// Communication API/ISOBUS/J1939-76/API/bds_isobus_initCnsrSdgDatabox
///This function initializes a J1939-76 consumer databox. The  J1939-76 messages can be sent only with  J1939-76 consumer databoxes.
///
///=======
/// Remarks:
///=======
/// + This function must be called during the configuration of the ISOBUS/J1939 and J1939-76 communication stack once for each J1939-76 consumer message.
/// + Before the consumer databoxes can be initialized with this function, the required number of receive databoxes has to be configured first with easyConfig tool or alternatively with function bds_isobus_registerCnsrSdgDataboxes.
/// + Each J1939-76 consumer databox requires an own data array or a data structure. The pointer to this data field is required for the initialization of a J1939-76 consumer databox. The received data then will be stored in this data field.
/// + The data array for the received data shall have length less than or equal to 8 (see parameter description below). 
/// + The execution time of the callback function should be short to be able to meet the time conditions within the ISOBUS/J1939 stack.
/// + If the same CAN bus is also used for further communication, ensure that the CAN IDs are uniquely assigned.
/// + The meaning of this function is similar to the ISOBUS/J1939 function bds_isobus_initRxDatabox.
/// + In addition to the ISOBUS/J1939 specifications, this function can be used for the reception of J1939-76 PDU1 format messages which are sent to the own network adddress as well as to other destination addresses.
/// + The definition of a destination address within PDU1 format PGNs is mandatory.
/// + Important: For the reception of PDU1 format messages to the own network address the PDU specific part (=Destination) of the PGN should be defined with the NULL address value (=0xFE) instead of the own address. Otherwise the own address within the RX databoxes may not match any more with the real own address after an address claiming.  
/// + The header file bds_bsw.h is included for enabling usage of defines.
///
///----------
/// FFI:
///----------
///This API can be used in trusted partitions only. See Freedom from Interference (FFI) concept for more details.
///
///
///Return value    																		Description
///==================================================================		  			===================================================================================================
///0: bds_isobus_sfty_noErr_E															Function executed without error
///3: bds_isobus_sfty_invldInstNum_E													Invalid ISOBUS/J1939 CA instance number
///7: bds_isobus_sfty_invldDataboxNum_E													Invalid databox number
///8: bds_isobus_sfty_invldPgn_E														Invalid PGN
///9: bds_isobus_sfty_invldPrio_E														Invalid priority
///10: bds_isobus_sfty_invldCyc_E														Invalid cycle time
///11: bds_isobus_sfty_invldOffs_E														Invalid offset time.
///12: bds_isobus_sfty_invldDataLen_E													Invalid data length
///13: bds_isobus_sfty_invldDataPtr_E													invalid pointer address
///14: bds_isobus_sfty_pgnPrioExists_E													Another databox with the same PGN and priority is already defined.
///15: bds_isobus_sfty_invldSrcAdr_E													Invalid Source Address
///16: bds_isobus_sfty_invldSct_E														Invalid SCT value
///17: bds_isobus_sfty_invldSrvt_E														Invalid SRVT value	
///19: bds_isobus_sfty_featNotEnad_E													API used without enabling J1939-76 feature in easyConfig
///20: bds_isobus_sfty_invldCbkAdr_E 													Callback function value NULL is invalid. Callback function is mandatory for J1939-76
///					  									
///==================================================================		   			===================================================================================================
///
///
///==================================================================		  			===================================================================================================
///Standard PGN	 								  										Data in Databox
///==================================================================		  			===================================================================================================
///Registered as "0xEEFF"																Receives only data which is broadcasted (PDU Specific part =0xFF).
///																						ex: bds_isobus_initCnsrSdgDatabox(1u, 1u, 0xEEFF, 0x10, 120, 50, 8, cnsrSDMdata_au8, NULL);
///																						It only receives the data which is brodcasted from source address 0x10.
///
///Registered "0xEE<own address>"														Receives data which is directed to the ECU by its own address (PDU Specific part=Destination).
///																						ex: bds_isobus_initCnsrSdgDatabox(1u, 1u, 0xEE04, 0x10, 120, 50, 8, cnsrSDMdata_au8, NULL);
///																						It only receives the data which is directed TO the ECU BY requesting with its own address(0x04).
///																					    Note: IF you initialize databox with "0xEEFE" you only receive data with whose PDU Specific part is Null(0xFE).
///==================================================================		   			===================================================================================================
///
///=======
///Code Example:
///=======
///============================================================================
///
/// PROGRAM Isobus_test
/// VAR_GLOBAL
///  cnsrMsg1Data_au8: ARRAY[1..8] OF USINT;
///
/// END_VAR
///	
/// 
/// VAR
///	   ISOBUS_SFTY_CNSR_BOXES_DU8: USINT :=35;
///    registerApiRetVal_e : bds_isobus_sfty_apiRetVal_te;    
///    initApi1RetVal_e : bds_isobus_sfty_apiRetVal_te;
///    isobus_sfty_cnsrSdgMsg_as: ARRAY[1..35] OF bds_isobus_cnsrSdgMsg_ts ;
///    instance_num:USINT:=1;
///
/// END_VAR
///
/// IF(Flag_u8=0) THEN
///
/// bds_can_init(BDS_CAN_3_D, BDS_BAUD_1000K_DU32); 	
///	bds_can_sendData(BDS_CAN_3_D, 16#999999, 1, 0,0);
///
/// registerApiRetVal_e := bds_isobus_registerCnsrSdgDataboxes(1, ADR(isobus_sfty_cnsrSdgMsg_as), ISOBUS_SFTY_CNSR_BOXES_DU8);
/// 
/// initApi1RetVal_e := bds_isobus_initCnsrSdgDatabox(1, 1, 16#4901, 16#10, 24, 100, 8, ADR(gvl.cnsrMsg1Data_au8), ADR(cnsrMsgCallback1));
///
/// bds_isobus_setCaName(instance_num,16#00,16#02,16#00,16#01,16#81,16#01,16#01,16#33,BDS_ISOBUS_OWN_SN_DU32);
///
/// bds_isobus_setCaName(instance_num,16#00,16#02,16#00,16#01,16#81,16#01,16#01,16#33,BDS_ISOBUS_OWN_SN_DU32);
/// 
/// retval5_u16:=bds_isobus_setCaAddr(instance_num,BDS_CAN_3_D,16#10);
///
/// bds_isobus_initComm(bds_can_Chnl_te.BDS_CAN_3_D, 50);
///
/// Flag_u8:=1;
/// 
/// END_IF
///
/// FUNCTION cnsrMsgCallback1 : UINT
/// VAR_INPUT	
///	data_length: POINTER TO BYTE;
///	data_pau8: POINTER TO BYTE ;
///	status_e : bds_isobus_sdgCnsrStatus_te;
/// END_VAR

/// VAR
///  i : INT;
///    cnsrCbk_rcvd_u32 : UDINT;
///    CbkSt_e : bds_isobus_sdgCnsrStatus_te;
///    CbkDataLen_u8 : POINTER TO BYTE:=0;
///	 data_au8: ARRAY [1..8] OF USINT:=[1,2];
/// END_VAR
///
/// cnsrCbk_rcvd_u32 := cnsrCbk_rcvd_u32 + 1;
/// CbkDataLen_u8 := data_length;
/// CbkSt_e := status_e;
///
/// FOR i := 0 TO 7 DO
/// gvl.cnsrMsg1Data_au8[i] := data_pau8[i];  // Dereference pointer to copy each element
/// END_FOR;
/// END
///============================================================================

{attribute 'external_name' := 'cmp_rts_bds_isobus_initCnsrSdgDatabox'}

FUNCTION bds_isobus_initCnsrSdgDatabox : bds_isobus_sfty_apiRetVal_te
VAR_INPUT
	///ISOBUS/J1939 instance number. This number identifies one instance of the ISOBUS/J1939 stack.
 	///
	///Value range: 1..n
	///n is the number of ISOBUS instances configured by easyConfig. 
	instanceNum_u8 : USINT;
	///Number of a J1939-76 producer databox.
	///
	///Value range: 1..n
	///n is the number of producer databoxes configured by easyConfig or alternatively with function bds_isobus_registerProdSdgDataboxes.
	sdgDataboxNum_u16 : UINT;
	///Parameter group number (PGN) of the SDM(Safety Data Message) to be sent with this databox.
	///
	///Value range: 0..0x3FFFF (18 bit) 
	///The lowest byte of the PGN contains for:
	/// + PDU1 format:  the destination address
	/// + PDU2 format:  the PDU extension
	pgn_u32 : UDINT;
	///Source address of the J1939-76 consumer from where the message has to be received.
	///
	///
	///Value range: 0x00..0xFD 
	src_u8 : USINT;
	///The maximum time interval in ms between two consecutive SDMs received.
	///
	///
	///Value Range: 10ms - 65000ms
	sct_u32 : UDINT;
	///The maximum time interval in ms between an SHM and SDM of an SDG received.
	///
	///
	///Value Range: 10ms - 65000ms
	srvt_u32 : UDINT;
	///Size of the data to be received. A J1939-76 consumer message data size must be less than or equal to 8 bytes.
	//
	///Value range: 1...8 bytes
	lenMax_u8 : USINT;
	///Pointer to a data array, in which the received data can be stored.
	/// The size of this array/structure has to be given within the previous parameter (lenMax_u8).
	///
	///It is neccessary to declare the data buffer array as a global variable.
	data_pau8: POINTER TO USINT;
	///Pointer to callback function of type bds_isobus_sdgCnsrCallback_tpf which will be called after reception and processing of a consumer SDG.
	func_pf: POINTER TO UINT;
END_VAR

END_FUNCTION

// Communication API/ISOBUS/J1939-76/API/bds_isobus_registerCnsrSdgDataboxes
///This function registers memory for J1939-76 safety extension consumer databoxes and therefore defines the maximal number of usable J1939-76 consumer databoxes per instance.
///
///=======
/// Remarks:
///=======
///		+ This function must be called once during the configuration of the ISOBUS/J1939 communication stack before bds_isobus_initComm.
/// 	+ After the execution of this function, each  J1939-76 consumer databox has to be initialized with bds_isobus_initCnsrSdgDatabox before using the databoxes.
/// 	+ The header file bds_bsw.h is included for enabling usage of defines.
/// 
///----------
/// FFI:
///----------
///
///This API can be used in trusted partitions only. See Freedom from Interference (FFI) concept for more details.
///	
///==================================================================		  			===================================================================================================
///Return value    								  									Description
///==================================================================		  			===================================================================================================
/// 0: bds_isobus_sfty_noErr_E 																Function executed without error
/// 1: bds_isobus_sfty_invldAdr_E															invalid address of databox (mem_pas)
/// 2: bds_isobus_sfty_ovlAdr_E                                                             Address overlaps with an already existing buffer.
/// 3: bds_isobus_sfty_invldInstNum_E                                                       Invalid CA instance number
///	6: bds_isobus_sfty_cfgNotAllwd_E                                                        Function must be called before bds_isobus_initComm, but it was called afterwards.																			-
/// 19: bds_isobus_sfty_featNotEnad_E                                                       API used without enabling J1939-76 feature in easyConfig
///
///
///==================================================================		   			===================================================================================================
///
/// Code Example:
///=======
///============================================================================
/// PROGRAM Isobus_test
/// VAR_GLOBAL
///  cnsrMsg1Data_au8: ARRAY[1..8] OF USINT;
///
/// END_VAR
///	
/// 
/// VAR
///	   ISOBUS_SFTY_CNSR_BOXES_DU8: USINT :=35;
///    registerApiRetVal_e : bds_isobus_sfty_apiRetVal_te;    
///    initApi1RetVal_e : bds_isobus_sfty_apiRetVal_te;
///    isobus_sfty_cnsrSdgMsg_as: ARRAY[1..35] OF bds_isobus_cnsrSdgMsg_ts ;
///    instance_num:USINT:=1;
///
/// END_VAR
///
/// IF(Flag_u8=0) THEN
///
/// bds_can_init(BDS_CAN_3_D, BDS_BAUD_1000K_DU32); 	
///	bds_can_sendData(BDS_CAN_3_D, 16#999999, 1, 0,0);
///
/// registerApiRetVal_e := bds_isobus_registerCnsrSdgDataboxes(1, ADR(isobus_sfty_cnsrSdgMsg_as), ISOBUS_SFTY_CNSR_BOXES_DU8);
/// 
/// initApi1RetVal_e := bds_isobus_initCnsrSdgDatabox(1, 1, 16#4901, 16#10, 24, 100, 8, ADR(gvl.cnsrMsg1Data_au8), ADR(cnsrMsgCallback1));
///
/// bds_isobus_setCaName(instance_num,16#00,16#02,16#00,16#01,16#81,16#01,16#01,16#33,BDS_ISOBUS_OWN_SN_DU32);
///
/// bds_isobus_setCaName(instance_num,16#00,16#02,16#00,16#01,16#81,16#01,16#01,16#33,BDS_ISOBUS_OWN_SN_DU32);
/// 
/// retval5_u16:=bds_isobus_setCaAddr(instance_num,BDS_CAN_3_D,16#10);
///
/// bds_isobus_initComm(bds_can_Chnl_te.BDS_CAN_3_D, 50);
///
/// Flag_u8:=1;
/// 
/// END_IF
///
/// FUNCTION cnsrMsgCallback1 : UINT
/// VAR_INPUT	
///	data_length: POINTER TO BYTE;
///	data_pau8: POINTER TO BYTE ;
///	status_e : bds_isobus_sdgCnsrStatus_te;
/// END_VAR

/// VAR
///  i : INT;
///    cnsrCbk_rcvd_u32 : UDINT;
///    CbkSt_e : bds_isobus_sdgCnsrStatus_te;
///    CbkDataLen_u8 : POINTER TO BYTE:=0;
///	 data_au8: ARRAY [1..8] OF USINT:=[1,2];
/// END_VAR
///
/// cnsrCbk_rcvd_u32 := cnsrCbk_rcvd_u32 + 1;
/// CbkDataLen_u8 := data_length;
/// CbkSt_e := status_e;
///
/// FOR i := 0 TO 7 DO
/// gvl.cnsrMsg1Data_au8[i] := data_pau8[i];  // Dereference pointer to copy each element
/// END_FOR;
/// END
///============================================================================


{attribute 'external_name' := 'cmp_rts_bds_isobus_registerCnsrSdgDataboxes'}
FUNCTION bds_isobus_registerCnsrSdgDataboxes : bds_isobus_sfty_apiRetVal_te
VAR_INPUT
	///ISOBUS/J1939 instance number. This number identifies one instance of the ISOBUS/J1939 stack.
	///
	///Value range: 1..n
	///n is the number of ISOBUS/J1939 instances configured in easyConfig. 
	instanceNum_u8 : USINT;
	///Pointer to an array of data type bds_isobus_cnsrSdgMsg_ts.
	///
	///Note:
	///The buffer will be managed by the C-API. The application has only to declare the buffer (memory space).It is necessary to declare the buffer array as a global variable.
	mem_pas : POINTER TO  bds_isobus_prodSdgMsg_ts;
	///Size of the array above, which corresponds to the number of usable J1939-76 consumer databoxes.
	numOfMsg_u16: UINT;
END_VAR

END_FUNCTION

// Communication API/ISOBUS/J1939-76/API/bds_isobus_registerProdSdgDataboxes
///This function registers memory for J1939-76 safety extension producer databoxes and therefore defines the maximal number of usable J1939-76 producer databoxes per instance.
///
///=======
/// Remarks:
///=======
///		+ This function must be called once during the configuration of the ISOBUS/J1939 communication stack before bds_isobus_initComm.
/// 	+ After the execution of this function, each J1939-76 producer databox has to be initialized with bds_isobus_initProdDatabox before using the databoxes.
///     + The header file bds_bsw.h is included for enabling usage of defines.
///
///----------
/// FFI:
///----------
///This API can be used in trusted partitions only. See Freedom from Interference (FFI) concept for more details.
///
///==================================================================		  			===================================================================================================
///Return value    								  									     Description
///==================================================================		  			===================================================================================================
///0: bds_isobus_sfty_noErr_E															Function executed without error
///1: bds_isobus_sfty_invldAdr_E														Invalid address of databox (*mem_pas)
///2: bds_isobus_sfty_ovlAdr_E															Address overlaps with an already existing buffer.
///3: bds_isobus_sfty_invldInstNum_E													invalid CA instance number.
///6: bds_isobus_sfty_cfgNotAllwd_E														Function must be called before bds_isobus_initComm, but it was called afterwards.
///19: bds_isobus_sfty_featNotEnad_E													API used without enabling J1939-76 feature in easyConfig
///
/// 
///==================================================================		   			===================================================================================================
///
/// Code Example:
///=======
///============================================================================
/// PROGRAM Isobus_test
/// VAR_GLOBAL
///  prodMsg2Data_au8: ARRAY[1..8] OF USINT:=[16#A,16#1,16#2,16#3,16#4,16#5,16#6,16#7];
///
/// END_VAR
///
/// VAR
///
///    registerApiRetVal_e : bds_isobus_sfty_apiRetVal_te;    
///    initApi1RetVal_e : bds_isobus_sfty_apiRetVal_te;
///    isobus_sfty_prodSdgMsg_as: ARRAY[1..34] OF bds_isobus_prodSdgMsg_ts  ;
///    instance_num:USINT:=1;
///
/// END_VAR
///
/// IF(Flag_u8=0) THEN
///
/// bds_can_init(BDS_CAN_3_D, BDS_BAUD_1000K_DU32); 	
///	bds_can_sendData(BDS_CAN_3_D, 16#999999, 1, 0,0);
///
/// registerApiRetVal_e := bds_isobus_registerProdSdgDataboxes(instance_num,ADR(isobus_sfty_prodSdgMsg_as), 35);
/// 
/// initApi1RetVal_e := bds_isobus_initProdSdgDatabox(instance_num,1,16#4410,6, 100 , 10 , 8 , ADR(gvl.prodMsg2Data_au8) ,ADR(ProdMsgCallback1));
///
/// bds_isobus_setCaName(instance_num,16#00,16#02,16#00,16#01,16#81,16#01,16#01,16#33,BDS_ISOBUS_OWN_SN_DU32);
///
/// bds_isobus_setCaName(instance_num,16#00,16#02,16#00,16#01,16#81,16#01,16#01,16#33,BDS_ISOBUS_OWN_SN_DU32);
/// 
/// retval5_u16:=bds_isobus_setCaAddr(instance_num,BDS_CAN_3_D,16#10);
///
/// bds_isobus_initComm(bds_can_Chnl_te.BDS_CAN_3_D, 50);
///
/// Flag_u8:=1;
/// 
/// END_IF
///
/// FUNCTION ProdMsgCallback1 : USINT
/// 
/// VAR_INPUT
/// data_length:POINTER TO BYTE;
/// data_pau8: POINTER TO BYTE;
/// END_VAR
///
/// data_pau8[0] := 16#07;
/// data_pau8[1] := 16#06;
/// data_pau8[2] := 16#05;
/// data_pau8[3] := 16#04;
/// data_pau8[4] := 16#03;
/// data_pau8[5] := 16#FF;
/// data_pau8[6] := 16#FF;
/// data_pau8[7] := 16#FF;
/// 
/// data_length[0]:=8;
///
/// END
///============================================================================
{attribute 'external_name' := 'cmp_rts_bds_isobus_registerProdSdgDataboxes'}
FUNCTION bds_isobus_registerProdSdgDataboxes : bds_isobus_sfty_apiRetVal_te
VAR_INPUT
	///ISOBUS/J1939 instance number. This number identifies one instance of the ISOBUS/J1939 stack.
	///
	///Value range: 1..n
	///n is the number of ISOBUS/J1939 instances configured in easyConfig. 
	instanceNum_u8 : USINT;
	///Pointer to an array of data type bds_isobus_prodSdgMsg_ts. 
	///
	///Note:
	///The buffer will be managed by the C-API. The application has only to declare the buffer (memory space).
	///It is necessary to declare the buffer array as a global variable.
	mem_pas : POINTER TO  bds_isobus_prodSdgMsg_ts;
	///Size of the array, which corresponds to the number of usable J1939-76 producer databoxes.  
	numOfMsg_u16: UINT;
END_VAR

END_FUNCTION

// Communication API/ISOBUS/J1939-76/API/bds_isobus_initProdSdgDatabox
///This function initializes a J1939-76 producer databox. The J1939-76 messages can be sent only with J1939-76 producer databoxes.
///=======
/// Remarks:
///=======
/// + This function must be called during the configuration of the ISOBUS/J1939 and J1939-76 communication stack once for each J1939-76 producer message.
/// + Before the producer databoxes can be initialized with this function, the required number of producer databoxes has to be configured first with easyConfig tool or alternatively with function bds_isobus_registerProdSdgDataboxes.
/// + Each J1939-76 producer databox requires an own data array or a data structure. The pointer to this data field is required for the initialization of a J1939-76 producer databox. The transmitted data will be taken from this data field.
/// + The data array for the transmitted data must have a length of less than or equal to 8 bytes (see parameter description below).
/// + The execution time of the callback function should be short to be able to meet the time conditions within the ISOBUS/J1939 stack. 
/// + If the same CAN bus is also used for further communication, ensure that the CAN IDs are uniquely assigned.
/// + The meaning of this function is similar to the ISOBUS/J1939 function bds_isobus_initTxDatabox.
/// + The header file bds_bsw.h is included for enabling usage of defines.

///----------
/// FFI:
///----------
///This API can be used in trusted partitions only. See Freedom from Interference (FFI) concept for more details.
///
///==================================================================		  			===================================================================================================
///Return value    								  									Description
///==================================================================		  			===================================================================================================
///0: bds_isobus_sfty_noErr_E                                                             Function executed without error
///3: bds_isobus_sfty_invldInstNum_E                                                      Invalid ISOBUS/J1939 CA instance number
///7: bds_isobus_sfty_invldDataboxNum_E                                                   invalid databox number
///8: bds_isobus_sfty_invldPgn_E                                                          Invalid PGN
///9: bds_isobus_sfty_invldPrio_E                                                         Invalid priority
///10: bds_isobus_sfty_invldCyc_E                                                         Invalid cycle time
///11: bds_isobus_sfty_invldOffs_E                                                        Invalid offset time.
///12: bds_isobus_sfty_invldDataLen_E                                                     Invalid data length. 
///13: bds_isobus_sfty_invldDataPtr_E                                                     Invalid pointer address
///14: bds_isobus_sfty_pgnPrioExists_E                                                    Another databox with the same PGN and priority is already defined.

///==================================================================		   			===================================================================================================
///
///=======
///Code Example:
///=======
///
/// PROGRAM Isobus_test
/// VAR_GLOBAL
///  prodMsg2Data_au8: ARRAY[1..8] OF USINT:=[16#A,16#1,16#2,16#3,16#4,16#5,16#6,16#7];
///
/// END_VAR
///
/// VAR
///
///    registerApiRetVal_e : bds_isobus_sfty_apiRetVal_te;    
///    initApi1RetVal_e : bds_isobus_sfty_apiRetVal_te;
///    isobus_sfty_prodSdgMsg_as: ARRAY[1..34] OF bds_isobus_prodSdgMsg_ts  ;
///    instance_num:USINT:=1;
///
/// END_VAR
///
/// IF(Flag_u8=0) THEN
///
/// bds_can_init(BDS_CAN_3_D, BDS_BAUD_1000K_DU32); 	
///	bds_can_sendData(BDS_CAN_3_D, 16#999999, 1, 0,0);
///
/// registerApiRetVal_e := bds_isobus_registerProdSdgDataboxes(instance_num,ADR(isobus_sfty_prodSdgMsg_as), 35);
/// 
/// initApi1RetVal_e := bds_isobus_initProdSdgDatabox(instance_num,1,16#4410,6, 100 , 10 , 8 , ADR(gvl.prodMsg2Data_au8) ,ADR(ProdMsgCallback1));
///
/// bds_isobus_setCaName(instance_num,16#00,16#02,16#00,16#01,16#81,16#01,16#01,16#33,BDS_ISOBUS_OWN_SN_DU32);
///
/// bds_isobus_setCaName(instance_num,16#00,16#02,16#00,16#01,16#81,16#01,16#01,16#33,BDS_ISOBUS_OWN_SN_DU32);
/// 
/// retval5_u16:=bds_isobus_setCaAddr(instance_num,BDS_CAN_3_D,16#10);
///
/// bds_isobus_initComm(bds_can_Chnl_te.BDS_CAN_3_D, 50);
///
/// Flag_u8:=1;
/// 
/// END_IF
///
///
/// FUNCTION ProdMsgCallback1 : USINT
/// 
/// VAR_INPUT
/// data_length:POINTER TO BYTE;
/// data_pau8: POINTER TO BYTE;
/// END_VAR
///
/// data_pau8[0] := 16#07;
/// data_pau8[1] := 16#06;
/// data_pau8[2] := 16#05;
/// data_pau8[3] := 16#04;
/// data_pau8[4] := 16#03;
/// data_pau8[5] := 16#FF;
/// data_pau8[6] := 16#FF;
/// data_pau8[7] := 16#FF;
/// 
/// data_length[0]:=8;
///
/// END
///============================================================================

{attribute 'external_name' := 'cmp_rts_bds_isobus_initProdSdgDatabox'}
FUNCTION bds_isobus_initProdSdgDatabox : bds_isobus_sfty_apiRetVal_te
VAR_INPUT
	///ISOBUS/J1939 instance number. This number identifies one instance of the ISOBUS/J1939 stack.
 	///
	///Value range: 1..n
	///n is the number of ISOBUS instances configured by easyConfig. 
	instanceNum_u8 : USINT;
	///Number of a J1939-76 producer databox.
	///
	///Value range: 1..n
	///n is the number of producer databoxes configured by easyConfig or alternatively with function bds_isobus_registerProdSdgDataboxes.
	sdgDataboxNum_u16 : UINT;
	///Parameter group number (PGN) of the SDM(Safety Data Message) to be sent with this databox.
	///
	///Value range: 0..0x3FFFF (18 bit) 
	///The lowest byte of the PGN contains for:
	/// + PDU1 format:  the destination address
	/// + PDU2 format:  the PDU extension
	pgn_u32 : UDINT;
	///Priority of the message to be sent.
	///
	///Value range: 0..7  (6 = default value according ISOBUS/J1939 specification)
	prio_u8 : USINT;
	/// This time (in ms) controls the cyclic transmission (or) fixed transmission of the J1939-76 Producer message from this J1939-76 producer databox.
	///The cycle time of a J1939-76 producer message must be greater than or equal to 10ms.
	///Cycle time value 0 is invalid.
	///Value range: 10..65000 [ms].
	cycle_u16 : UINT;
	///The first transmission cycle of a J1939-76 producer message can be shortened by this offset time (in ms). 
	///This can be used to prevent CAN bus overload, if several messages have to be sent with the same cycle time.
	///With an offset = 0 the first message will be sent after the cycle time.
	///
	///Value range: 0.. (cycle_u16 - 1) [ms]
	offset_u16 : UINT;
	///Size of the data to be transmitted in bytes. A J1939-76 producer message data size must be less than or equal to 8.
	/// 
	///Value range: 1...8 bytes
	lenMax_u8 : USINT;
	///Pointer to a data array, from which the data is taken for transmission.  
	///The size of this array has to be given within the previous parameter (lenMax_u8).
	///
	///It is necessary to declare the data array as a global variable.
	data_pau8: POINTER TO USINT;
	///Pointer to callback function of type bds_isobus_sdgProdCallback_tpf which will be called by
	///BSW FOR data update BY ASW before transmission OF a producer SDG.
	func_pf: POINTER TO USINT;
END_VAR

END_FUNCTION

// Diagnostics API/UDS/API/Vehicle Identification Number(VIN) APIs/bds_uds_setVin
///This function sets the Vehicle Identification Number(VIN) of the ECU.
///
///=======
///Additional Info: + The Vehicle Identification Number(VIN) configured in the ECU is mapped to the DID 0xF190.
///					+ By default, the VIN has a value of B0DASMACH1NE00001.
///=======
///
///=======
/// Remarks: 
///=======
///			+ This function must be called from OsIniProc().
/// 		+ The header file bds_bsw.h is included for enabling usage of defines.
///
///-----------
///
/// FFI:
///----------
///This API can be used in trusted partitions only. See Freedom from Interference (FFI) concept for more details.
///
///
///==================================================================		  			===================================================================================================
///Return value    								  									Description
///==================================================================		  			===================================================================================================
///bds_udsCmn_ok_E																		API call successful.
///bds_udsCmn_invldPrm_E																API call invalid because of an invalid parameter.
///bds_udsCmn_outOfRng_E																Out of range, the array size should be less than or equal to 17 bytes.
///bds_udsCmn_notAvl_E																	not available (e.g. busy, called to early in init, system is in a mode that it cannot measure, etc)
///==================================================================		   			===================================================================================================
///
///=======
///Code Example:
///=======
///PROGRAM Vin_test
/// VAR
/// setVin_pau8:ARRAY[0..16] OF USINT:=[16#54,16#45 ,16#53 ,16#54 ,16#56 ,16#49 ,16#4E ,16#42 ,16#4F ,16#44 ,16#41 ,16#53 ,16#31 ,16#32 ,16#33 ,16#34 ,16#35];
/// flag_1:USINT;
/// retval_e:  bds_udsCmn_statusApi_te;
/// END_VAR
///
/// IF(flag_1=0) THEN
/// retval_e:=bds_uds_setVin(ADR(setVin_pau8),17);
/// flag_1:=1;
/// END_IF
//=============================================
{attribute 'external_name' := 'cmp_rts_bds_uds_setVin'}
FUNCTION bds_uds_setVin : bds_udsCmn_statusApi_te
VAR_INPUT
	//Pointer to set/configure the VIN data which is mapped to the DID 0xF190.
	data_pau8: POINTER TO USINT;
	//Size of the Vehicle Identification Number in bytes.
	size_u8: USINT;
END_VAR

END_FUNCTION

// Diagnostics API/UDS/API/Vehicle Identification Number(VIN) APIs/bds_uds_getVin
///This function reads the Vehicle Identification Number(VIN) of the ECU.
///
///=======
///Additional Info: + The Vehicle Identification Number(VIN) configured in the ECU is mapped to the DID 0xF190.
///					+ By default, the VIN has a value of B0DASMACH1NE00001.
///=======
///
///=======
/// Remarks: 
///=======
/// 		+ The header file bds_bsw.h is included for enabling usage of defines.
///
///-----------
///
/// FFI:
///----------
///This API can be used in trusted partitions only. See Freedom from Interference (FFI) concept for more details.
///
///
///==================================================================		  			===================================================================================================
///Return value    								  									Description
///==================================================================		  			===================================================================================================
///bds_udsCmn_ok_E																		API call successful.
///bds_udsCmn_invldPrm_E																API call invalid because of an invalid parameter.
///bds_udsCmn_outOfRng_E																Out of range, the array size should be less than or equal to 17 bytes.
///
///==================================================================		   			===================================================================================================
///
///=======
///Code Example:
///=======
///PROGRAM Vin_test
/// VAR
/// getVin_pau8:ARRAY[0..16] OF USINT;
/// 
/// retval_e:  bds_udsCmn_statusApi_te;
/// END_VAR
///
/// 
/// retval_e:=bds_uds_setVin(ADR(setVin_pau8),17);
/// 
/// retval_e:=bds_uds_getVin(ADR(getVin_pau8),APPL_VIN_SIZE_DU8);
//=============================================
{attribute 'external_name' := 'cmp_rts_bds_uds_getVin'}
FUNCTION bds_uds_getVin : bds_udsCmn_statusApi_te
VAR_INPUT
	//Pointer to set/configure the VIN data which is mapped to the DID 0xF190.
	data_pau8: POINTER TO USINT;
	//Size of the Vehicle Identification Number in bytes.
	size_u8: USINT;
END_VAR

END_FUNCTION

// Diagnostics API/UDS/API/Vehicle Identification Number(VIN) APIs/bds_uds_registerVinCallback
///This function registers the read and write callbacks for the DID 0xF190 used for the Vehicle Identification Number (VIN).
///
///=======
///Additional Info: + The Vehicle Identification Number(VIN) configured in the ECU is mapped to the DID 0xF190.
///					+ By default, the VIN has a value of B0DASMACH1NE00001.
///=======
///=======
/// Remarks: 
///=======
/// 		+ The header file bds_bsw.h is included for enabling usage of defines.
///
///-----------
/// FFI:
///----------
///This API can be used in trusted partitions only. See Freedom from Interference (FFI) concept for more details.
///
///
///==================================================================		  			===================================================================================================
///Return value    								  									Description
///==================================================================		  			===================================================================================================
///bds_udsCmn_ok_E																		API call successful.
///bds_udsCmn_invldPrm_E																API call invalid because of an invalid parameter.
///bds_udsCmn_outOfRng_E																Out of range, the array size should be less than or equal to 17 bytes.
///bds_udsCmn_notAvl_E																	not available (e.g. busy, called to early in init, system is in a mode that it cannot measure, etc)
///==================================================================		   			===================================================================================================
///
///=======
///Code Example:
///=======
/// VAR_GLOBAL
///	 read_data:ARRAY[0..16] OF USINT:=[16#54,16#45 ,16#53 ,16#54 ,16#56 ,16#49 ,16#4E ,16#42 ,16#4F ,16#44 ,16#41 ,16#53 ,16#31 ,16#32 ,16#33 ,16#34 ,16#35];
/// END_VAR
///
/// PROGRAM Vin_test
/// VAR
///
/// retval_e:  bds_udsCmn_statusApi_te;
/// flag_1:USINT;
///
/// END_VAR
/// 
/// IF(flag_1=0) THEN 
/// retval_e:=bds_uds_registerVinCallback(ADR(vinReadCallbackfunc), ADR(vinWriteCallbackfunc));
/// flag_1:=1;
/// END_IF
/// 
/// FUNCTION vinReadCallbackfunc : USINT
/// VAR_INPUT
///	Data:POINTER TO USINT;
///END_VAR
///
/// VAR
///	i : USINT;
///	readVinCntr : INT;
///	data_au8 : ARRAY[0..7] OF USINT:=[2,4];
/// END_VAR
/// 
/// FOR i:= 0 TO 16 DO
///	Data[i]:=gvl.read[i];
/// END_FOR
/// 
/// readVinCntr:= readVinCntr+1;
/// 
/// FUNCTION vinWriteCallbackfunc : USINT
/// VAR_INPUT
///	Data:POINTER TO USINT;
///	errorCode_pu8:POINTER TO USINT;	
///END_VAR
///
/// VAR
///	writeVinCntr : INT;
///	data_au8 : ARRAY[0..7] OF USINT:=[1,2];
///	i:USINT:=0;
/// END_VAR
/// 
/// FOR i:= 0 TO 16 DO
///	Data[i]:=gvl.read[i];
/// END_FOR
/// writeVinCntr:=writeVinCntr+1;
///
/// 
///=============================	
{attribute 'external_name' := 'cmp_rts_bds_uds_registerVinCallback'}
FUNCTION bds_uds_registerVinCallback : bds_udsCmn_statusApi_te
VAR_INPUT
	//Pointer to a callback function which is called if a VIN is read through DID 0xF190 read.
	funcRead_pf: POINTER TO USINT;
	//Pointer to a callback function which is called if a VIN is written through DID 0xF190 write.
	funcWrite_pf: POINTER TO USINT;
END_VAR

END_FUNCTION

// Communication API/CAN/CAN-FD legacy/API/bds_can_fd_registerRxCallback
///This function allows for the registration of a callback function for a CAN-FD supported CAN channel. The callback function is triggered when a CAN-FD message is received in the registered CAN channel.
///
///=======
/// Remarks:
///=======
///There are some alternatives for handling incoming CAN-FD messages (combinations are allowed):
///- Receive buffer which has to be defined with easyConfig. Function bds_can_fd_getData has to be used in order to get received messages.
///- Callback function which has to be registered with function described. 
///- Receive databoxes which have to be configured with easyConfig. Each receive databox has to be initialized with function bds_can_fd_initRxDatabox. Function bds_can_fd_getDatabox has to be used in order to get a message from a receive databox.
///Registering of this callback function is optional.
///This callback function will not be called for messages for which a receive databox was defined with function bds_can_fd_initRxDatabox.
///This function call is allowed only in initialization task.
///This callback function must be defined within the application program.
///The CAN-FD callback functions registered with this API are executed in core-0.
///The header file bds_cmn_bsw.h is included for enabling usage of defines.
///
///----------
/// FFI:
///----------
///This API can be used in trusted partitions.See Freedom from Interference (FFI) concept for more details.
///
///----------
/// WARNING:
///----------
///The callback function has a higher priority than user tasks.
///It is recommended to use this function only for code that can be executed fast, e.g. to save data. 
///Adding more code in callback function implies that runtime of the function increases, which may influence user tasks.
///
///==================================================================		  			===================================================================================================
///Return value    								  										Description
///==================================================================		  			===================================================================================================
///0 - bds_can_fd_ok_E																	API call successful, CAN-FD Receive callback is registered successfully
///14 - bds_can_fd_invldChnl_E                                                          Invalid CAN channel called
///60 - bds_can_fd_invldAddr_E                                                          Invalid address (CAN-FD Receive callback function address pointed wrong)
///99 - bds_can_fd_cfgNotAllowed_E                                                      Configuration is not allowed.
///                                                                                     Note: Configuration has to be made only during initialization e.g., in OsIniProc().
///100 - bds_can_fd_paramChnl3Err_E                                                     CAN-FD is not supported on CAN_3.
///==================================================================		   			===================================================================================================
///
///=======
///Code Example:
///=======
///PROGRAM Test_for_T3_can_fd
///VAR
/// flag_u8:USINT:=0;
///END_VAR
///
///IF (flag_u8 = 0) THEN
///bds_can_fd_registerRxCallback(bds_can_chnl_te.BDS_CAN_1_D, ADR(can_2_fd_RxCallback));
///flag_u8:=1;
///
///FUNCTION can_2_fd_RxCallback : UINT
///VAR_INPUT
///	format_u8 : USINT;
///	id_u32 : UDINT;
///	numBytes_u8 : USINT;
///	data_pau8 : POINTER TO USINT;
///END_VAR

/// store received message data and evaluate them outside of this callback!
///============================================================================                                
{attribute 'external_name' := 'cmp_rts_bds_can_fd_registerRxCallback'}
FUNCTION bds_can_fd_registerRxCallback : bds_can_fd_St_te
VAR_INPUT
	//Indicates the CAN channel.
	//Possible values :
	//BDS_CAN_1_D(0)
	//BDS_CAN_2_D(1)
	//BDS_CAN_4_D(3)
	chnl_e:bds_can_Chnl_te;
	//Pointer to a callback function of data type bds_can_RxCallback_tpf which is called if a CAN message was received.
	func_pf : POINTER TO UINT;
END_VAR

END_FUNCTION

// Communication API/CAN/CAN-FD legacy/API/bds_can_fd_initRxDatabox
///This function initializes a CAN-FD receive databox for a specified CAN channel.By initialization, it means that the CAN-FD receive databox is assigned with the following parameters:
///- Databox number
///- CAN ID
///- CAN ID format
///- Number of bytes of data
///- CAN-FD Receive Databox data buffer
///- Databox buffer length
///- Callback function time
///
///=======
/// Remarks:
///=======
/// The use of CAN-FD receive databoxes is optional!
/// The number of required CAN-FD receive databoxes must be defined in easyConfig before using this function.
/// Each CAN-FD receive databox has to be initialized before it can be used.
/// The CAN-FD callback functions registered with this API are executed in core-0.
/// The header file bds_cmn_bsw.h is included for enabling usage of defines.
///
///----------
/// FFI:
///----------
///This API can be used in trusted partitions.See Freedom from Interference (FFI) concept for more details.
///
///==================================================================		  			===================================================================================================
///Return value    								  										Description
///==================================================================		  			===================================================================================================
///0: bds_can_fd_ok_E                                                                   Function is called without errors. Receive databox was initialized successfully.
///9: bds_can_fd_invldDataBoxNbr_E                                                      Invalid CAN-FD databox number.
///14: bds_can_fd_invldChnl_E                                                           Unknown CAN channel.
///15: bds_can_fd_invldId_E                                                             Invalid CAN identifier.
///16: bds_can_fd_invldFormat_E                                                         Invalid message format.
///17: bds_can_fd_invldNumBytes_E                                                       Invalid number of data bytes.
///55: bds_can_fd_ovlpAddr_E                                                            Buffer overlaps with buffer registered already.
///60: bds_can_fd_invldAddr_E                                                           NA.
///61: bds_can_fd_rxDataboxBufLenZero_E                                                 Invalid address (parameter buf_pas).Buffer length is zero.
///63: bds_can_fd_errDataboxIdExist_E                                                   A databox with this identifier is initialised already.The new initialization will be not accepted.
///100 - bds_can_fd_paramChnl3Err_E                                                     CAN-FD not supported for CAN_3
///
///==================================================================		   			===================================================================================================
///
///=======
///Code Example:
///=======
///PROGRAM Test_for_T3_can_fd
///VAR_GLOBAL
///can_2_fd_RxDatabox_2_Buf_as : ARRAY[0..7] OF bds_can_fd_DataboxData_ts;
///testRxBox_as:ARRAY[0..7] OF bds_can_fd_RxDatabox_ts;
///VAR_END
///
///VAR
///CAN_2_FD_RX_DATABOX_2_BUF_LEN_DU8 : USINT :=1;
///bds_can_fd_St_te apiStatusRxBoxReg_e;
///bds_can_fd_St_te apiStatusRxBoxInit_e;
///bds_can_fd_St_te apiStatusRxBoxRcv_e;
/// flag_u8 : USINT:=0;
///END_VAR
///
///IF(flag_u8 = 0) THEN 
///apiStatusRxBoxReg_e:=bds_can_fd_registerRxDataboxes(bds_can_chnl_te.BDS_CAN_1_D, ADR(GVL.testRxBox_as[0]), 10);
///
///apiStatusRxBoxInit_e:=bds_can_fd_initRxDatabox(bds_can_chnl_te.BDS_CAN_1_D,1,16#701,BDS_CAN_STD_DU8,8,
///                ADR(GVL.can_2_fd_RxDatabox_2_Buf_as),CAN_2_FD_RX_DATABOX_2_BUF_LEN_DU8,ADR(can_2_fd_RxDatabox_2_Callback));
///
///bds_can_initxt(bds_can_chnl_te.BDS_CAN_1_D, BDS_BAUD_250K_DU32, 81, BDS_BAUD_2000K_DU32);
///
///flag_u8:=1;
///
///FUNCTION can_2_fd_RxDatabox_2_Callback 
///VAR_INPUT
///
///END_VAR
///VAR
///	DataboxData_au8 : ARRAY[0..7] OF USINT;
///	DataboxNumBytes_u8 : USINT;
///	data_pau8 : ARRAY[0..2] OF USINT:=[1,2,3];
///END_VAR
///
///bds_can_fd_getDatabox(bds_can_chnl_te.BDS_CAN_1_D, 1, ADR(DataboxData_au8), DataboxNumBytes_u8);
///============================================================================
{attribute 'external_name' := 'cmp_rts_bds_can_fd_initRxDatabox'}
FUNCTION bds_can_fd_initRxDatabox : bds_can_fd_St_te
VAR_INPUT
	//Indicates the CAN channel.
	//Possible values :
	//BDS_CAN_1_D(0)
	//BDS_CAN_2_D(1)
	//BDS_CAN_4_D(3)
	chnl_e : bds_can_Chnl_te;
	//Receive databox number.
	//Each receive databox is numbered separately for each CAN channel.Value range: 1 .. n.
	//n is the number of databoxes configured by easyConfig. 
	databoxNum_u16 : UINT;
	//Identifier of CAN message.Value range:
	//16#000 .. 0x7FF (11-bit standard format)
	//16#00000000 .. 0x1FFFFFFF (29-bit extented format)
	id_u32 : UDINT;
	//Indicates the format of the CAN-FD message.Value range:
	//BDS_CAN_STD_DU8  (11-bit standard format)
	//BDS_CAN_EXD_DU8  (29-bit extented format)
	format_u8 : USINT;
	//Number of bytes which can be received at maximum.Value range: 0 .. 64
	numBytes_u8 : USINT;
	//Pointer to array of data type bds_can_fd_DataboxData_ts.
	//Note:The buffer will be managed by C-API. The application has only to declare the buffer (memory space). 
    //It is recommended to declare the buffer array in a local function with attribute "static".
	buf_pas : POINTER TO bds_can_fd_DataboxData_ts;
	//Length of buffer array (that means number of CAN-FD messages).At least a buffer for 1 message is required.
	buf_len_u16 : UINT;
	//Pointer to a callback function to receive a new message
	callback_pf : POINTER TO UINT;
END_VAR

END_FUNCTION

// Communication API/CAN/CAN-FD legacy/API/bds_can_fd_registerRxDataboxes
///This API registers memory for CAN-FD receive databoxes of a CAN channel.
///
///=======
/// Remarks:
///=======
///Usage of this API is optional.
///This API shall be used if: 
///- User needs to configure and use more CAN-FD receive databoxes (maximum number of receive databoxes which shall be configured in easyConfig is 40 and minimum of 1 transmit databox shall be configured).
///- User doesn't need to configure CAN-FD receive databoxes in easyConfig.
///Using this API will overwrite the number of CAN-FD receive databoxes used in easyConfig.
///This API shall be called only in initialization task.
///The header file bds_cmn_bsw.h is included for enabling usage of defines.
///
///=======
/// INFO:
///=======
///This API shall be preferred to be used only when user needs to configure more than 40 CAN-FD Receive Databoxes.
///Memory usage information:
///- bds_can_fd_RxDatabox_ts mem_as[1] - 24 bytes = Memory reserved for one CAN-FD Receive Databox.Additionally, 
///1. Number of bytes required for initialization = bds_can_fd_DataboxData_ts rxBox1_as[1] = 65 bytes for buffer size 1 (CAN-FD Receive Databox buffer size)
///2. Databox data = 64 bytes of data
///Hence it is advised to declare databox handle buffer keeping memory usage into account.Sample usage is seen in How to configure CAN-FD legacy using Transmit, Receive Databoxes.
///
///----------
/// FFI:
///----------
///This API can be used in trusted partitions.See Freedom from Interference (FFI) concept for more details.
///
///==================================================================		  			===================================================================================================
///Return value    								  										Description
///==================================================================		  			===================================================================================================
///0 - bds_can_fd_ok_E																	API call successful.
///14 - bds_can_fd_invldChnl_E                                                          Invalid CAN channel because invalid CAN channel passed.
///60 - bds_can_fd_invldAddr_E                                                          Invalid address, e.g., because NULL pointer was passed for pointer to structure of bds_can_fd_RxDatabox_ts.
///64 - bds_can_fd_prevRegdDataboxMoreThanCurrent_E                                     Number of databoxes registered is greater than previously registered number of databoxes.
///65 - bds_can_fd_invldCfgDatabox_E                                                    Invalid number of databoxes used for configuration, e.g., number of configured databoxes = 0.
///99 - bds_can_fd_cfgNotAllowed_E                                                      Configuration of Rx databoxes not allowed, i.e., API call happened in ASW Initialization task.
///100 - bds_can_fd_paramChnl3Err_E                                                     CAN-FD not supported in CAN_3.
///
///==================================================================		   			===================================================================================================
///
///=======
///Code Example:
///=======
///PROGRAM Test_for_T3_can_fd
///VAR_GLOBAL
///can_2_fd_RxDatabox_2_Buf_as : ARRAY[0..7] OF bds_can_fd_DataboxData_ts;
///testRxBox_as:ARRAY[0..7] OF bds_can_fd_RxDatabox_ts;
///VAR_END
///
///VAR
///CAN_2_FD_RX_DATABOX_2_BUF_LEN_DU8 : USINT :=1;
///bds_can_fd_St_te apiStatusRxBoxReg_e;
///bds_can_fd_St_te apiStatusRxBoxInit_e;
///bds_can_fd_St_te apiStatusRxBoxRcv_e;
///flag_uu8:USINT:=0;
///END_VAR
///
///IF(flag_u8 = 0 ) THEN
///apiStatusRxBoxReg_e:= bds_can_fd_registerRxDataboxes(bds_can_chnl_te.BDS_CAN_1_D, ADR(GVL.testRxBox_as[0]), 10);
///
///apiStatusRxBoxInit_e:= bds_can_fd_initRxDatabox(bds_can_chnl_te.BDS_CAN_1_D,1,16#701,BDS_CAN_STD_DU8,8,
///                ADR(GVL.can_2_fd_RxDatabox_2_Buf_as),CAN_2_FD_RX_DATABOX_2_BUF_LEN_DU8,ADR(can_2_fd_RxDatabox_2_Callback));
///
///bds_can_initxt(bds_can_chnl_te.BDS_CAN_1_D, BDS_BAUD_250K_DU32, 81, BDS_BAUD_2000K_DU32);
///flag_u8:=1;
///
///
///FUNCTION can_2_fd_RxDatabox_2_Callback 
///VAR_INPUT
///
///END_VAR
///VAR
///	DataboxData_au8 : ARRAY[0..7] OF USINT;
///	DataboxNumBytes_u8 : USINT;
///	data_pau8 : ARRAY[0..2] OF USINT:=[1,2,3];
///END_VAR
///
///bds_can_fd_getDatabox(bds_can_chnl_te.BDS_CAN_1_D, 1, ADR(DataboxData_au8), DataboxNumBytes_u8);
///============================================================================
{attribute 'external_name' := 'cmp_rts_bds_can_fd_registerRxDataboxes'}
FUNCTION bds_can_fd_registerRxDataboxes : bds_can_fd_St_te
VAR_INPUT
	//Indicates the CAN channel.
	//Possible values :
	//BDS_CAN_1_D(0)
	//BDS_CAN_2_D(1)
	//BDS_CAN_4_D(3)
	chnl_e : bds_can_Chnl_te;
	//Pointer to a structure of type bds_can_fd_RxDatabox_ts.Note: This buffer will be used for Receive databox handling. 
	mem_pas: POINTER TO bds_can_fd_RxDatabox_ts;
	//Number of receive databoxes
    num_u16: UINT; 
END_VAR

END_FUNCTION

// Communication API/CAN/CAN-FD legacy/API/bds_can_fd_getDatabox
///This API gets a message from the specified CAN-FD receive databox of the specified CAN channel.
///- If the databox was initialized with a buffer length = 1 then the last received message will be read from the databox buffer.
///- If the databox was initialized with a buffer length > 1 then the oldest message will be read from the databox buffer.
///
///=======
/// Remarks:
///=======
/// The specified receive databox has to be initialized by bds_can_fd_initRxDatabox before using this function.
/// The number of required receive databoxes must be defined by easyConfig before using this function.
/// The header file bds_cmn_bsw.h is included for enabling usage of defines.
///
///----------
/// FFI:
///----------
///This API can be used in trusted partitions. For untrusted partitions use bds_can_fd_getDatabox_ffi. See Freedom from Interference (FFI) concept for more details.
///
///==================================================================		  			===================================================================================================
///Return value    								  										Description
///==================================================================		  			===================================================================================================
///0: bds_can_fd_ok_E                                                                   Function is called without errors. Message data returned in data_pau8 are valid.
///5: bds_can_fd_errFfi_E                                                               Invalid Access to FFI variant API call.
///9: bds_can_fd_invldDataBoxNbr_E                                                      Invalid transmit databox number.
///14: bds_can_fd_invldChnl_E                                                           Unknown CAN channel.
///30: bds_can_fd_rxBufOvfl_E                                                           Receive buffer overflow. At least one message is lost. Message data returned in msg_s are valid.
///31: bds_can_fd_rxBufEmpty_E                                                          Receive buffer is empty. Message data returned in msg_s are invalid.
///60: bds_can_fd_invldAddr_E                                                           Invalid address (parameter msg_s).
///62: bds_can_fd_dataBoxNoInit_E                                                       Databox is not initialized.
///100 - bds_can_fd_paramChnl3Err_E                                                     CAN-FD not supported for CAN_3
///
///==================================================================		   			===================================================================================================
///
///=======
///Code Example:
///=======
///PROGRAM Test_for_T3_can_fd
///VAR_GLOBAL
///can_2_fd_RxDatabox_2_Buf_as : ARRAY[0..7] OF bds_can_fd_DataboxData_ts;
///testRxBox_as:ARRAY[0..7] OF bds_can_fd_RxDatabox_ts;
///VAR_END
///
///VAR
///CAN_2_FD_RX_DATABOX_2_BUF_LEN_DU8 : USINT :=1;
///bds_can_fd_St_te apiStatusRxBoxReg_e;
///bds_can_fd_St_te apiStatusRxBoxInit_e;
///bds_can_fd_St_te apiStatusRxBoxRcv_e;
///END_VAR
///
///IF(flag_u8 = 0) THEN
///bds_can_fd_registerRxDataboxes(bds_can_chnl_te.BDS_CAN_1_D, ADR(GVL.testRxBox_as[0]), 10);
///
///bds_can_fd_initRxDatabox(bds_can_chnl_te.BDS_CAN_1_D,1,16#701,BDS_CAN_STD_DU8,8,
///                ADR(GVL.can_2_fd_RxDatabox_2_Buf_as),CAN_2_FD_RX_DATABOX_2_BUF_LEN_DU8,ADR(can_2_fd_RxDatabox_2_Callback));
///
///bds_can_initxt(bds_can_chnl_te.BDS_CAN_1_D, BDS_BAUD_250K_DU32, 81, BDS_BAUD_2000K_DU32);
///
///flag_u8:=1;
///
///FUNCTION can_2_fd_RxDatabox_2_Callback 
///VAR_INPUT
///
///END_VAR
///VAR
///	DataboxData_au8 : ARRAY[0..7] OF USINT;
///	DataboxNumBytes_u8 : USINT;
///	data_pau8 : ARRAY[0..2] OF USINT:=[1,2,3];
///END_VAR
///
///bds_can_fd_getDatabox(bds_can_chnl_te.BDS_CAN_1_D, 1, ADR(DataboxData_au8), DataboxNumBytes_u8);
///============================================================================
{attribute 'external_name' := 'cmp_rts_bds_can_fd_getDatabox'}
FUNCTION bds_can_fd_getDatabox : bds_can_fd_St_te
VAR_INPUT
	//Indicates the CAN channel.
	//Possible values :
	//BDS_CAN_1_D(0)
	//BDS_CAN_2_D(1)
	//BDS_CAN_4_D(3)
	chnl_e : bds_can_Chnl_te;
	//CAN-FD Receive databox number.
	//Each receive databox is numbered separately for each CAN channel.
	//n is the number of databoxes configured by easyConfig. 
	databoxNum_u16 : UINT;
	//Pointer to data array.The oldest data received by the configured databox is copied to this address. 
    data_pau8 :POINTER TO USINT;
	//Number of bytes which are copied to data array data_pau8.
	numBytes_pu8 :POINTER TO USINT;
END_VAR

END_FUNCTION

// Communication API/CAN/CAN_FD_FFI_API/bds_can_fd_getDatabox_ffi
{attribute 'external_name' := 'cmp_rts_bds_can_fd_getDatabox_ffi'}
FUNCTION bds_can_fd_getDatabox_ffi : bds_can_fd_St_te
VAR_INPUT
	//Indicates the CAN channel.
	//Possible values :
	//BDS_CAN_1_D(0)
	//BDS_CAN_2_D(1)
	//BDS_CAN_4_D(3)
	chnl_e : bds_can_Chnl_te;
	//CAN-FD Receive databox number.
	//Each receive databox is numbered separately for each CAN channel.
	//n is the number of databoxes configured by easyConfig. 
	databoxNum_u16 : UINT;
	//Pointer to data array.The oldest data received by the configured databox is copied to this address. 
    data_pau8 :POINTER TO USINT;
	//Number of bytes which are copied to data array data_pau8.
	numBytes_pu8 :POINTER TO USINT;
END_VAR

END_FUNCTION

// Communication API/CAN/CAN-FD legacy/API/bds_can_fd_registerTxDataboxes
///This API registers memory for CAN-FD receive databoxes of a CAN channel.
///
///=======
/// Remarks:
///=======
///Usage of this API is optional.
///This API shall be used if: 
///- User needs to configure and use more CAN-FD receive databoxes (maximum number of receive databoxes which shall be configured in easyConfig is 40 and minimum of 1 transmit databox shall be configured).
///- User doesn't need to configure CAN-FD receive databoxes in easyConfig.
///Using this API will overwrite the number of CAN-FD receive databoxes used in easyConfig.
///This API shall be called only in initialization task.
///The header file bds_cmn_bsw.h is included for enabling usage of defines.
///
///=======
/// INFO:
///=======
///This API shall be preferred to be used only when user needs to configure more than 40 CAN-FD Receive Databoxes.
///Memory usage information:
///- bds_can_fd_TxDatabox_ts mem_as[1] - 72 bytes = Memory reserved for one Transmit DataboxAdditionally, 
///1. Number of bytes required for transmission = 64 bytes during API call (for Transmit Databox array)
///Hence it is advised to declare databox handle buffer keeping memory usage into account.Sample usage is seen in How to configure CAN-FD legacy using Transmit, Receive Databoxes.
///
///----------
/// FFI:
///----------
///This API can be used in trusted partitions.See Freedom from Interference (FFI) concept for more details.
///
///==================================================================		  			===================================================================================================
///Return value    								  										Description
///==================================================================		  			===================================================================================================
///0 - bds_can_fd_ok_E																	API call successful.
///14 - bds_can_fd_invldChnl_E                                                          Invalid CAN channel because invalid CAN channel passed.
///60 - bds_can_fd_invldAddr_E                                                          Invalid address, e.g., because NULL pointer was passed for pointer to structure of bds_can_fd_TxDatabox_ts.
///64 - bds_can_fd_prevRegdDataboxMoreThanCurrent_E                                     Number of databoxes registered is greater than previously registered number of databoxes.
///65 - bds_can_fd_invldCfgDatabox_E                                                    Invalid number of databoxes used for configuration, e.g., number of configured databoxes = 0.
///99 - bds_can_fd_cfgNotAllowed_E                                                      Configuration of Tx databoxes not allowed, i.e., API call happened in ASW Initialization task.
///100 - bds_can_fd_paramChnl3Err_E                                                     CAN-FD not supported in CAN_3.
///
///==================================================================		   			===================================================================================================
///
///=======
///Code Example:
///=======
///PROGRAM Test_for_T3_can_fd
///VAR_GLOBAL
///testRxBox_as:ARRAY[0..7] OF bds_can_fd_RxDatabox_ts;
///VAR_END
///
///VAR
///data_pau8 : ARRAY[0..63] OF USINT:=[1,2,3,4,5,6,7,8];
/// flag_u8: USINT:=0
///VAR_END
///
///IF(flag_u8 = 0) THEN
///bds_can_fd_registerTxDataboxes(bds_can_chnl_te.BDS_CAN_1_D, ADR(testTxBox_as), 10);
///
///bds_can_fd_initTxDatabox(bds_can_chnl_te.BDS_CAN_1_D, 1, 16#34, BDS_CAN_STD_DU8);
///
///flag_u8:=1;
///
///bds_can_fd_sendDatabox(bds_can_chnl_te.BDS_CAN_1_D,1,64,ADR(data_pau8));
///============================================================================
{attribute 'external_name' := 'cmp_rts_bds_can_fd_registerTxDataboxes'}
FUNCTION bds_can_fd_registerTxDataboxes : bds_can_fd_St_te
VAR_INPUT
	//Indicates the CAN channel.
	//Possible values :
	//BDS_CAN_1_D(0)
	//BDS_CAN_2_D(1)
	//BDS_CAN_4_D(3)
	chnl_e : bds_can_Chnl_te;
	//Pointer to a structure of type bds_can_fd_RxDatabox_ts.Note: This buffer will be used for Receive databox handling. 
	mem_pas: POINTER TO bds_can_fd_TxDatabox_ts;
	//Number of receive databoxes
    num_u16: UINT;
END_VAR

END_FUNCTION

// Communication API/CAN/CAN-FD legacy/API/bds_can_fd_initTxDatabox
///This function initializes, i.e., set a dedicated CAN ID and format (set databox parameters) to a CAN-FD transmit databox.
///
///=======
/// Remarks:
///=======
/// The use of transmit databoxes is optional.
/// The transmit databoxes must be defined in easyConfig before using this function.
/// Each transmit databox has to be initialized before it can be used.
/// If a transmit databox is initialized already it can be re-inititalized again (initialization of existing databox with different parameters such as ID, format). 
/// The header file bds_cmn_bsw.h is included for enabling usage of defines.
///
///----------
/// FFI:
///----------
///This API can be used in trusted partitions.See Freedom from Interference (FFI) concept for more details.
///
///==================================================================		  			===================================================================================================
///Return value    								  										Description
///==================================================================		  			===================================================================================================
///0: bds_can_fd_ok_E                                                                   Function is called without errors. Receive databox was initialized successfully.
///9: bds_can_fd_invldDataBoxNbr_E                                                      Invalid transmit databox number.
///14: bds_can_fd_invldChnl_E                                                           Unknown CAN channel.
///15: bds_can_fd_invldId_E                                                             Invalid CAN identifier.
///16: bds_can_fd_invldFormat_E                                                         Invalid message format.
///100 - bds_can_fd_paramChnl3Err_E                                                     CAN-FD not supported for CAN_3
///
///==================================================================		   			===================================================================================================
///
///=======
///Code Example:
///=======
///PROGRAM Test_for_T3_can_fd
///VAR_GLOBAL
///testRxBox_as:ARRAY[0..7] OF bds_can_fd_RxDatabox_ts;
///VAR_END
///
///VAR
///data_pau8 : ARRAY[0..63] OF USINT:=[1,2,3,4,5,6,7,8];
/// flag_u8: USINT:=0
///VAR_END
///
///IF(flag_u8 = 0) THEN
///bds_can_fd_registerTxDataboxes(bds_can_chnl_te.BDS_CAN_1_D, ADR(testTxBox_as), 10);
///
///bds_can_fd_initTxDatabox(bds_can_chnl_te.BDS_CAN_1_D, 1, 16#34, BDS_CAN_STD_DU8);
///
///flag_u8:=1;
///
///bds_can_fd_sendDatabox(bds_can_chnl_te.BDS_CAN_1_D,1,64,ADR(data_pau8));
///============================================================================
{attribute 'external_name' := 'cmp_rts_bds_can_fd_initTxDatabox'}
FUNCTION bds_can_fd_initTxDatabox : bds_can_fd_St_te
VAR_INPUT
	//Indicates the CAN channel.
	//Possible values :
	//BDS_CAN_1_D(0)
	//BDS_CAN_2_D(1)
	//BDS_CAN_4_D(3)
	chnl_e : bds_can_Chnl_te;
	//Transmit databox number.
	//Each transmit databox is numbered separately for each CAN channel.Value range: 1 .. n.
	//n is the number of databoxes configured by easyConfig. 
	databoxNum_u16 : UINT;
	//Identifier of CAN message.Value range:
	//16#000 .. 0x7FF (11-bit standard format)
	//16#00000000 .. 0x1FFFFFFF (29-bit extented format)
	id_u32 : UDINT;
	//Indicates the format of the CAN-FD message.Value range:
	//BDS_CAN_STD_DU8  (11-bit standard format)
	//BDS_CAN_EXD_DU8  (29-bit extented format)
	format_u8 : USINT;	
END_VAR

END_FUNCTION

// Communication API/CAN/CAN-FD legacy/API/bds_can_fd_sendDatabox
///This API sends a CAN-FD message via a transmit databox.
///
///=======
/// Remarks:
///=======
/// The number of required transmit databoxes must be defined by easyConfig.
/// The specified transmit databox has to be initialized by bds_can_fd_initTxDatabox before using this function.
/// A transmit databox buffers only the actual message.
/// A message in a transmit databox (which was not sent) can be overwritten by a new order. No error will occur!
/// Function bds_can_fd_isTxDataboxFree can be used in order to check whether a transmit databox is free again.
/// Messages in transmit data boxes will be sent before messages in transmit buffer (bds_can_fd_sendData).
/// The time interval for sending the messages can be defined with the function bds_can_fd_setTxDelay.
/// The header file bds_cmn_bsw.h is included for enabling usage of defines.
///
///----------
/// FFI:
///----------
///This API can be used in trusted partitions. For untrusted partitions use bds_can_fd_getDatabox_ffi. See Freedom from Interference (FFI) concept for more details.
///
///==================================================================		  			===================================================================================================
///Return value    								  										Description
///==================================================================		  			===================================================================================================
///0: bds_can_fd_ok_E                                                                   Function is called without errors. Message data returned in data_pau8 are valid.
///5: bds_can_fd_errFfi_E                                                               Invalid Access to FFI variant API call.
///9: bds_can_fd_invldDataBoxNbr_E                                                      Invalid transmit databox number.
///14: bds_can_fd_invldChnl_E                                                           Unknown CAN channel.
///17: bds_can_fd_invldNumBytes_E                                                       Invalid number of data bytes.
///60: bds_can_fd_invldAddr_E                                                           Invalid address (parameter msg_s).
///62: bds_can_fd_dataBoxNoInit_E                                                       Transmit databox is not initialized.
///100 - bds_can_fd_paramChnl3Err_E                                                     CAN-FD not supported for CAN_3
///
///==================================================================		   			===================================================================================================
///
///=======
///Code Example:
///=======
///PROGRAM Test_for_T3_can_fd
///VAR_GLOBAL
///testRxBox_as:ARRAY[0..7] OF bds_can_fd_RxDatabox_ts;
///VAR_END
///
///VAR
///data_pau8 : ARRAY[0..63] OF USINT:=[1,2,3,4,5,6,7,8];
/// flag_u8: USINT:=0
///VAR_END
///
///IF(flag_u8 = 0) THEN
///bds_can_fd_registerTxDataboxes(bds_can_chnl_te.BDS_CAN_1_D, ADR(testTxBox_as), 10);
///
///bds_can_fd_initTxDatabox(bds_can_chnl_te.BDS_CAN_1_D, 1, 16#34, BDS_CAN_STD_DU8);
///
///flag_u8:=1;
///
///bds_can_fd_sendDatabox(bds_can_chnl_te.BDS_CAN_1_D,1,64,ADR(data_pau8));
///============================================================================
{attribute 'external_name' := 'cmp_rts_bds_can_fd_sendDatabox'}
FUNCTION bds_can_fd_sendDatabox : bds_can_fd_St_te
VAR_INPUT
	//Indicates the CAN channel.
	//Possible values :
	//BDS_CAN_1_D(0)
	//BDS_CAN_2_D(1)
	//BDS_CAN_4_D(3)
	chnl_e : bds_can_Chnl_te;
	//Transmit databox number.
	//Each transmit databox is numbered separately for each CAN channel.Value range: 1 .. n.
	//n is the number of databoxes configured by easyConfig. 
	itxdataboxNum_u16 : UINT;
	//Number of bytes to be sent.Value range: 0 .. 64
	numBytes_pu8 : USINT;
	//Pointer to array of data bytes. The number of bytes is contained in parameter numBytes_u8. 
    //A NULL pointer is allowed if number of data bytes (parameter numBytes_u8) is zero. 
    data_pau8 :POINTER TO USINT;
END_VAR

END_FUNCTION

// Communication API/CAN/CAN-FD legacy/API/bds_can_fd_isTxDataboxFree
///This function checks whether a CAN-FD transmit databox is free again. 
///A transmit databox is free again if it was possible to send the last CAN-FD message via the bus.
///
///=======
/// Remarks:
///=======
///The use of transmit databoxes is optional.
///The transmit databoxes of that CAN channel has to be defined by easyConfig tool and that transmit databox has to be initialised by bds_can_fd_initTxDatabox before using this function.
///This function can be used to prevent overwriting of a message that has not yet been sent in a send databox, by checking whether the previous message was actually sent before writing the new message to the databox.
///The time it takes for a databox to become available for sending again depends greatly on the baud rate and the bus load.
///The header file bds_cmn_bsw.h is included for enabling usage of defines.
///
///----------
/// FFI:
///----------
///This API can be used in trusted partitions. For untrusted partitions use  bds_can_fd_isTxDataboxFree_ffi.. See Freedom from Interference (FFI) concept for more details.
///
///==================================================================		  			===================================================================================================
///Return value    								  										Description
///==================================================================		  			===================================================================================================
///0: bds_can_fd_ok_E                                                                   No error. Databox is empty.
///1: bds_can_fd_txDataboxNotEmpty_E                                                    No error. Databox is not empty.
///5: bds_can_fd_errFfi_E                                                               Invalid Access to FFI variant API call.
///9: bds_can_fd_invldDataBoxNbr_E                                                      Invalid transmit databox number.
///14: bds_can_fd_invldChnl_E                                                           Unknown CAN channel.
///62: bds_can_fd_dataBoxNoInit_E                                                       Databox is not initialized.
///100 - bds_can_fd_paramChnl3Err_E                                                     CAN-FD not supported for CAN_3
///
///==================================================================		   			===================================================================================================
///=======
///Code Example:
///===============
///PROGRAM Test_for_T3_can_fd
///VAR_GLOBAL
///testRxBox_as:ARRAY[0..7] OF bds_can_fd_RxDatabox_ts;
///VAR_END
///
///VAR
///data_pau8 : ARRAY[0..63] OF USINT:=[1,2,3,4,5,6,7,8];
/// flag_u8: USINT:=0
///VAR_END
///
///IF(flag_u8 = 0) THEN
///bds_can_fd_registerTxDataboxes(bds_can_chnl_te.BDS_CAN_1_D, ADR(testTxBox_as), 10);
///
///bds_can_fd_initTxDatabox(bds_can_chnl_te.BDS_CAN_1_D, 1, 16#34, BDS_CAN_STD_DU8);
///
///flag_u8:=1;
///
///bds_can_fd_isTxDataboxFree(bds_can_chnl_te.BDS_CAN_1_D, 1);
///===========================================================
{attribute 'external_name' := 'cmp_rts_bds_can_fd_isTxDataboxFree'}
FUNCTION bds_can_fd_isTxDataboxFree : bds_can_fd_St_te
VAR_INPUT
	//Indicates the CAN channel.
	//Possible values :
	//BDS_CAN_1_D(0)
	//BDS_CAN_2_D(1)
	//BDS_CAN_4_D(3)
	chnl_e : bds_can_Chnl_te;
	//Transmit databox number.
    //Each transmit databox is numbered separately for each CAN channel.Value range: 1 .. n.
	//n is the number of databoxes configured by easyConfig. 
	txDataboxNum_u16 : UINT;
END_VAR

END_FUNCTION

// Communication API/CAN/CAN_FD_FFI_API/bds_can_fd_isTxDataboxFree_ffi
{attribute 'external_name' := 'cmp_rts_bds_can_fd_isTxDataboxFree_ffi'}
FUNCTION bds_can_fd_isTxDataboxFree_ffi : bds_can_fd_St_te
VAR_INPUT
	//Indicates the CAN channel.
	//Possible values :
	//BDS_CAN_1_D(0)
	//BDS_CAN_2_D(1)
	//BDS_CAN_4_D(3)
	chnl_e : bds_can_Chnl_te;
	//Transmit databox number.
    //Each transmit databox is numbered separately for each CAN channel.Value range: 1 .. n.
	//n is the number of databoxes configured by easyConfig. 
	txDataboxNum_u16 : UINT;
END_VAR

END_FUNCTION

// Communication API/CAN/CAN-FD legacy/API/bds_can_fd_setTxDelay
///The bds_can_fd_setTxDelay function can be used to define an optional delay time for sending CAN-FD messages for a CAN-FD supported CAN channel.
///Without executing this function the default delay time = 0 is used.
///A delay time > 0 should be only specified, if another controller is not able to receive the CAN-FD messages with full speed.
///
///=======
/// Remarks:
///=======
///Only messages which are sent with the functions bds_can_fd_sendDatabox, bds_can_fd_sendData and all messages of ISOBUS module will be delayed.
///For each CAN channel another delay time can be specified.
///Signal based CAN messages, XCP and UDS messages are not impacted by this function.
///If an error occurs during execution of this function, the actual delay time will be not modified.
///The header file bds_cmn_bsw.h is included for enabling usage of defines.
///
///----------
/// FFI:
///----------
///This API can be used in trusted partitions only. See Freedom from Interference (FFI) concept for more details.
///
///==================================================================		  			===================================================================================================
///Return value    								  										Description
///==================================================================		  			===================================================================================================
///0: bds_can_fd_ok_E                                                                   Function is called without errors.
///14: bds_can_fd_invldChnl_E                                                           Unknown CAN channel.
///100 : bds_can_fd_paramChnl3Err_E                                                     CAN-FD not supported for CAN_3
///
///==================================================================		   			===================================================================================================
///==============
/// Code Example
///==================
///PROGRAM Test_for_T3_can_fd
///VAR
///flag_u8:USINT:=0;
///data_pau8 : ARRAY[0..7] OF USINT:=[1,2,3,4,5,6,7,8];
///data_pau8_1 : ARRAY[0..7] OF USINT:=[63,62,61,60,59,58,57,56];
///END_VAR
///
///IF(flag_u8 = 0) THEN
///bds_can_fd_setTxDelay(BDS_CAN_2_D, 10);
///
///END_IF
///
///bds_can_fd_sendData(bds_can_chnl_te.BDS_CAN_1_D, 16#356, BDS_CAN_STD_DU8, 8, ADR(data_pau8));
///bds_can_fd_sendData(bds_can_chnl_te.BDS_CAN_1_D, 16#456, BDS_CAN_STD_DU8, 8, ADR(data_pau8_1));
///=======================================================
{attribute 'external_name' := 'cmp_rts_bds_can_fd_setTxDelay'}
FUNCTION bds_can_fd_setTxDelay : bds_can_fd_St_te
VAR_INPUT
	//Indicates the CAN channel.
	//Possible values :
	//BDS_CAN_1_D(0)
	//BDS_CAN_2_D(1)
	//BDS_CAN_4_D(3)
	chnl_e : bds_can_Chnl_te;
	//Minimum delay time in ms between two sent CAN-FD messages.Value range: 0 .. 65535.
 	//0 = no delay time, means that the can messages will be sent as fast as possible.
	time_u16 : UINT;
END_VAR

END_FUNCTION

// Communication API/CAN/CAN_FD_FFI_API/bds_can_fd_getRxBufStatus_ffi
{attribute 'external_name' := 'cmp_rts_bds_can_fd_getRxBufStatus_ffi'}
FUNCTION bds_can_fd_getRxBufStatus_ffi : DINT
VAR_INPUT
	//Indicates the CAN channel.
	//Possible values :
	// + BDS_CAN_1_D(0)
	// + BDS_CAN_2_D(1)
	// + BDS_CAN_4_D(3)
	chnl_e:bds_can_Chnl_te;
END_VAR

END_FUNCTION

// Communication API/CAN/CAN_FD_FFI_API/bds_can_fd_sendData_ffi
{attribute 'external_name' := 'cmp_rts_bds_can_fd_sendData_ffi'}
FUNCTION bds_can_fd_sendData_ffi : bds_can_fd_St_te
VAR_INPUT
	//Indicates the CAN channel.
	//Possible values :
	// + BDS_CAN_1_D(0)
	// + BDS_CAN_2_D(1)
	// + BDS_CAN_4_D(3)
	chnl_e: bds_can_Chnl_te; 
    //Identifier of CAN-FD message.
	//Value range:
	//0x000 .. 0x7FF (11-bit standard format .. 0x1FFFFFFF (29-BIT extented format
	id_u32: UDINT;
	//Indicates the format of the CAN-FD message.
	//Value range:
	//BDS_CAN_STD_DU8  (11-bit standard format)
	//BDS_CAN_EXD_DU8  (29-bit extented format)
 	format_u8 : USINT;
	//Number of bytes to be sent.
	//
	//Value range: 1 .. 64
	numBytes_u8: USINT;
	//Pointer to array of data bytes. The number of bytes is contained in parameter numBytes_u8.
	//A NULL pointer is allowed if number of data bytes (parameter numBytes_u8) is zero. 
	data_pau8: POINTER TO USINT;
END_VAR

END_FUNCTION

// Communication API/CAN/CAN_FD_FFI_API/bds_can_fd_getTxBufStatus_ffi
{attribute 'external_name' := 'cmp_rts_bds_can_fd_getTxBufStatus_ffi'}
FUNCTION bds_can_fd_getTxBufStatus_ffi : DINT
VAR_INPUT
	//Indicates the CAN channel.
	//Possible values :
	//BDS_CAN_1_D(0)
	//BDS_CAN_2_D(1)
	//BDS_CAN_4_D(3)
	chnl_e: bds_can_Chnl_te;
END_VAR

END_FUNCTION

// Communication API/CAN/CAN_FD_FFI_API/bds_can_fd_getData_ffi
{attribute 'external_name' := 'cmp_rts_bds_can_fd_getData_ffi'}
FUNCTION bds_can_fd_getData_ffi : bds_can_fd_St_te
VAR_INPUT
	//Indicates the CAN channel.
	//Possible values :
	//BDS_CAN_1_D(0)
	//BDS_CAN_2_D(1)
	//BDS_CAN_4_D(3)
	chnl_e:bds_can_Chnl_te;
	//Pointer to the message data of type bds_can_fd_Message_ts.
	msg_s: POINTER TO bds_can_fd_Message_ts;
END_VAR

END_FUNCTION

// Communication API/CAN/CAN_FD_FFI_API/bds_can_fd_isTxChannelFree_ffi
{attribute 'external_name' := 'cmp_rts_bds_can_fd_isTxChannelFree_ffi'}
FUNCTION bds_can_fd_isTxChannelFree_ffi : UINT
VAR_INPUT
	//Indicates the CAN channel.
	//Possible values :
	//BDS_CAN_1_D(0)
	//BDS_CAN_2_D(1)
	//BDS_CAN_4_D(3)
	chnl_e: bds_can_Chnl_te;
END_VAR

END_FUNCTION

// Communication API/CAN/CAN_FD_FFI_API/bds_can_fd_sendDatabox_ffi
{attribute 'external_name' := 'cmp_rts_bds_can_fd_sendDatabox_ffi'}
FUNCTION bds_can_fd_sendDatabox_ffi : bds_can_fd_St_te
VAR_INPUT
	//Indicates the CAN channel.
	//Possible values :
	//BDS_CAN_1_D(0)
	//BDS_CAN_2_D(1)
	//BDS_CAN_4_D(3)
	chnl_e : bds_can_Chnl_te;
	//Transmit databox number.
	//Each transmit databox is numbered separately for each CAN channel.Value range: 1 .. n.
	//n is the number of databoxes configured by easyConfig. 
	itxdataboxNum_u16 : UINT;
	//Number of bytes to be sent.Value range: 0 .. 64
	numBytes_pu8 : USINT;
	//Pointer to array of data bytes. The number of bytes is contained in parameter numBytes_u8. 
    //A NULL pointer is allowed if number of data bytes (parameter numBytes_u8) is zero. 
    data_pau8 :POINTER TO USINT;
END_VAR

END_FUNCTION

// Communication API/ISOBUS/API/bds_isobus_registerCaAddrTable
///This function registers the ISOBUS address info table for the specified ISOBUS instance.
///The address info table is a structure array of type bds_isobus_caAddrInfoTbl_ts which shall be declared in RC Application software and is registered to RC BSW through this function.
///The size of the structure array shall be decided based on the maximum possible number of CAs in the ISOBUS/J1939 network.
///
///=======
/// Remarks:
///=======
/// This function must be called once during the configuration of the ISOBUS communication stack before bds_isobus_initComm.
/// Maximum size of structure array is 255 (i.e noOfEntry_u8 <=255) since ISOBUS/J1939 supports only upto 253 CAs in the network.
/// ISOBUS lib will not store its own instance address in the ISOBUS address info table. It is anyway available via API bds_isobus_getCaAddr.
///
///----------
/// FFI:
///----------
///This API can be used in trusted partitions only. See Freedom from Interference (FFI) concept for more details.
///
///==================================================================		  			===================================================================================================
///Return value    								  										Description
///==================================================================		  			===================================================================================================
/// RBR_ISOBUS_RC_NO_ERRORS_DU16                                                        Function executed without any errors, address info table registered successfully.                                                                      
/// RBR_ISOBUS_RC_CFG_NOTALLOWED_DU16                                                   Function must be called before bds_isobus_initComm, but it was called afterward's.
/// RBR_ISOBUS_RC_INV_INST_NUM_DU16                                                     Invalid ISOBUS instance number.
/// RBR_ISOBUS_RC_OVERLAP_ADDR_DU16                                                     structure array pointed by addrTableMem_pas overlaps with an already existing variable/array registered for other functions.
/// RBR_ISOBUS_RC_INVALID_ADDR_DU16                                                     structure array pointed by addrTableMem_pas is NULL
///==================================================================		   			===================================================================================================
///
///=======
///Code Example:
///=======
///PROGRAM Test_for_isobus
///VAR
///	flag_u8 :USINT:=0;
///	APPL_ISOBUS_ADDRESSINFOTBL_DU8 : USINT :=10;
///	isobus_caAddrInfoTbl_as:ARRAY[0..9] OF bds_isobus_caAddrInfoTbl_ts;
/// ret_u16 : UDINT;
///END_VAR
///
///
///IF( flag_u8 = 0 ) THEN
///ret_u16:=bds_isobus_registerCaAddrTable(1,ADR(isobus_caAddrInfoTbl_as[0]),APPL_ISOBUS_ADDRESSINFOTBL_DU8);
///
///bds_isobus_initComm(bds_can_Chnl_te.BDS_CAN_3_D, 50);
///flag_u8:=1
///
///END_IF
///============================================================================
{attribute 'external_name' := 'cmp_rts_bds_isobus_registerCaAddrTable'}
FUNCTION bds_isobus_registerCaAddrTable : UINT
VAR_INPUT CONSTANT
	//ISOBUS instance number. This number identifies one instance of the ISOBUS stack.
    //Value range: 1..n
	//n is the total number of ISOBUS instances configured by easyConfig or bds_isobus_registerInstances() API. 
	instanceNum_u8 : USINT;
	//Pointer to the structure array of address info table of type bds_isobus_caAddrInfoTbl_ts
	addrTableMem_pas : POINTER TO bds_isobus_caAddrInfoTbl_ts;
	//Size of the structure array pointed by addrTableMem_pas.Value range: 1..255
    noOfEntry_u8 : USINT;
END_VAR

END_FUNCTION

// Communication API/ISOBUS/API/bds_isobus_registerCaAddrInfoCbk
///This function registers a callback for the specified ISOBUS instance to handle events related to the reception of ISOBUS address claim messages and updates to the ISOBUS address info table. 
///The callback function is of type bds_isobus_caAddrInfoCallback_tpf and is triggered for the following events, specified by bds_isobus_caAddrCbEventType_te:
///
///Address claim message received without table update: This occurs when an address claim message is received, but no updates are made to the address info table.
///This can happen if the table is not registered or is full, preventing new entries. This event is indicated by bds_isobus_addrClaimMsgRcv_E.
///
///Address table entry updated: This occurs when an address claim message is received and the address table is updated with a new address.  
///This happens when the received CA name is already present in the table.This event is indicated by bds_isobus_caTbleAddressUpdate_E.
///
///New entry created in address table: This occurs when an address claim message is received and a new entry of CA name and address is created in the address table.
///This happens when the received CA name is not already present in the table. This event is indicated by bds_isobus_caTbleNewEntry_E.
///
///=======
/// Remarks:
///=======
/// This function must be called once during the configuration of the ISOBUS communication stack before bds_isobus_initComm.
/// Based on the change in address, application software can reconfigure the databox in the callback function registered through this  function.
/// The callback function can be used independent of ISOBUS address info table feature. i,e. to indicate only reception of address claim message.
///----------
/// FFI:
///----------
///This API can be used in trusted partitions only. See Freedom from Interference (FFI) concept for more details.
///
///==================================================================		  			===================================================================================================
///Return value    								  										Description
///==================================================================		  			===================================================================================================
/// RBR_ISOBUS_RC_NO_ERRORS_DU16                                                        Function executed without any errors, callback is registered successfully.                                                                      
/// RBR_ISOBUS_RC_CFG_NOTALLOWED_DU16                                                   Function must be called before bds_isobus_initComm, but it was called afterward's.
/// RBR_ISOBUS_RC_INV_INST_NUM_DU16                                                     Invalid ISOBUS instance number.
/// RBR_ISOBUS_RC_INVALID_ADDR_DU16                                                     function pointer pointed by func_pf is NULL
///==================================================================		   			===================================================================================================
///
///=======
///Code Example:
///=======
///PROGRAM Test_for_isobus
///VAR
///	flag_u8 :USINT:=0;
/// ret_u16 : UDINT;
///END_VAR
///
///
///IF( flag_u8 = 0 ) THEN
///bds_isobus_registerCaAddrInfoCbk(1,ADR(appl_isobus_addrclmcallback));
///
///bds_isobus_initComm(bds_can_Chnl_te.BDS_CAN_3_D, 50);
///flag_u8:=1
///
///END_IF
///
///FUNCTION appl_isobus_addrclmcallback 
///VAR_INPUT
///	eventType_e : bds_isobus_caAddrCbEventType_te;
///	newClaimAddr : USINT;
///	caName_pu8 : POINTER TO USINT;
///END_VAR
///
///VAR
///	i:USINT;
///	data_pau8:ARRAY[0..7]OF USINT;
///	valueToSend : USINT:=16#02;
///END_VAR
///
///caName_pu8 := ADR(valueToSend);
///============================================================================
{attribute 'external_name' := 'cmp_rts_bds_isobus_registerCaAddrInfoCbk'}
FUNCTION bds_isobus_registerCaAddrInfoCbk : UINT
VAR_INPUT CONSTANT
	//ISOBUS instance number. This number identifies one instance of the ISOBUS stack.
    //Value range: 1..n
	//n is the total number of ISOBUS instances configured by easyConfig or bds_isobus_registerInstances() API
	instanceNum_u8 : USINT;
	//pointer to callback function
	addClaimInfoFunc_pf :POINTER TO UINT;
END_VAR

END_FUNCTION

// Communication API/ISOBUS/API/bds_isobus_getCaAddrByName
///This function returns the address associated with a specified ISOBUS CA Name for a given ISOBUS instance. 
///The function performs the following steps:
///- Address Lookup: Searches the ISOBUS Address Info table for an entry matching the provided CA Name
///- Address Retrieval: If a match is found, returns the address mapped to the CA Name. If no match is found, returns an invalid address (0xFE).
///
///=======
/// Remarks:
///=======
/// This function can be called in any cyclic tasks.
/// This function returns 0xFE for invalid ISOBUS instance or if ISOBUS Address Info table was not registered through bds_isobus_registerCaAddrTable function.
///----------
/// FFI:
///----------
///This API can be used in trusted partitions only. See Freedom from Interference (FFI) concept for more details.
///
///==================================================================		  			===================================================================================================
///Return value    								  										Description
///==================================================================		  			===================================================================================================
///0 .. 253                                                                             valid CA address for a given CA name
///254                                                                                  Null Address, because function was executed with an error.
///==================================================================		   			===================================================================================================
///
///=======
///Code Example:
///=======
///PROGRAM Test_for_isobus
///VAR
///	flag_u8 :USINT:=0;
///	APPL_ISOBUS_ADDRESSINFOTBL_DU8 : USINT :=10;
///	isobus_caAddrInfoTbl_as:ARRAY[0..9] OF bds_isobus_caAddrInfoTbl_ts;
/// ret_u16 : UDINT;
///END_VAR
///
///VAR_GLOBAL
///testCAname_au8:ARRAY[0..7]OF USINT:=[16#04,16#00,16#60,16#06,16#09,16#81,16#02,16#20];
///VAR_END

///IF( flag_u8 = 0 ) THEN
///ret_u16:=bds_isobus_registerCaAddrTable(1,ADR(isobus_caAddrInfoTbl_as[0]),APPL_ISOBUS_ADDRESSINFOTBL_DU8);
///
///bds_isobus_initComm(bds_can_Chnl_te.BDS_CAN_3_D, 50);
///flag_u8:=1
///
///END_IF
///
///bds_isobus_getCaAddrByName(APPL_ISOBUS_INSTANCE_1,ADR(GVL.testCAName[0]));
///============================================================================
{attribute 'external_name' := 'cmp_rts_bds_isobus_getCaAddrByName'}
FUNCTION bds_isobus_getCaAddrByName : USINT
VAR_INPUT CONSTANT
	//ISOBUS instance number. This number identifies one instance of the ISOBUS stack.
    //Value range: 1..n
	//n is the total number of ISOBUS instances configured by easyConfig or bds_isobus_registerInstances() API
	instanceNum_u8 : USINT;
	//Name of ISOBUS CA for which address needs to be fetched.
	caName_pu8 : POINTER TO USINT;
END_VAR

END_FUNCTION

// Communication API/ISOBUS/API/bds_isobus_getAddressInfoTblRecordSize
///This function will return the number of valid entries in the ISOBUS address info table. The valid entry in a address info table is a CA name and its address.
///The return value 0 indicate no entry in the ISOBUS address info table 
///
///=======
/// Remarks:
///=======
/// This function can be called in any cyclic tasks.
/// This function returns 0 for invalid ISOBUS instance or if ISOBUS Address Info table was not registered through bds_isobus_registerCaAddrTable function.
///----------
/// FFI:
///----------
///This API can be used in trusted partitions only. See Freedom from Interference (FFI) concept for more details.
///
///==================================================================		  			===================================================================================================
///Return value    								  										Description
///==================================================================		  			===================================================================================================
///0                                                                                     no valid entries in ISOBUS address info table or function executed with errors
///1..253                                                                                number of valied entries in ISOBUS address table
///==================================================================		   			===================================================================================================
///
///=======
///Code Example:
///=======
/// PROGRAM Test_for_isobus
///VAR
///	flag_u8 :USINT:=0;
///	APPL_ISOBUS_ADDRESSINFOTBL_DU8 : USINT :=10;
///	isobus_caAddrInfoTbl_as:ARRAY[0..9] OF bds_isobus_caAddrInfoTbl_ts;
/// ret_u16 : UDINT;
///END_VAR
///

///IF( flag_u8 = 0 ) THEN
///ret_u16:=bds_isobus_registerCaAddrTable(1,ADR(isobus_caAddrInfoTbl_as[0]),APPL_ISOBUS_ADDRESSINFOTBL_DU8);
///
///bds_isobus_initComm(bds_can_Chnl_te.BDS_CAN_3_D, 50);
///flag_u8:=1
///
///END_IF
///
///bds_isobus_getAddressInfoTblRecordSize(1);
///============================================================================
{attribute 'external_name' := 'cmp_rts_bds_isobus_getAddressInfoTblRecordSize'}
FUNCTION bds_isobus_getAddressInfoTblRecordSize : USINT
VAR_INPUT CONSTANT
	//ISOBUS instance number. This number identifies one instance of the ISOBUS stack.
    //Value range: 1..n
	//n is the total number of ISOBUS instances configured by easyConfig or bds_isobus_registerInstances() API
	instanceNum_u8 : USINT;
END_VAR

END_FUNCTION

// Diagnostics API/UDS/API/bds_uds_getActiveService
///This function gets the active UDS service running in the server/ECU.
///
///=======
/// Remarks:
///=======
/// By default, no UDS service will be running on the server/ECU until a UDS service request is made by the tester.
///	The header file bds_cmn_bsw.h is included for enabling usage of defines.
/// The API can be used in the Read DID callbacks to differentiate between UDS service requests for the 0x22 (Read Data by Identifier) and 0x2F (Input Output Control by Identifier) services. 
/// Refer to the sample code provided in the Integration of IOCBI in ASW for a detailed example.
///
///----------
/// FFI:
///----------
///This API can be used in trusted partitions only. See Freedom from Interference (FFI) concept for more details.
///
///==================================================================		  			===================================================================================================
///Return value    								  							            Description
///==================================================================		  			===================================================================================================
///bds_uds_getActiveService_ts															The return structure containing the status of API function call and the Service Identifier (SID) value.
///
///==================================================================		   			===================================================================================================
///
///=======
///Code Example:
///=======
///============================================================================
{attribute 'external_name' := 'cmp_rts_bds_uds_getActiveService'}
FUNCTION bds_uds_getActiveService : bds_uds_getActiveService_ts
VAR_INPUT
	// No parameters
END_VAR

END_FUNCTION

// System API/SYS/API/bds_sysSm_getCfg
///This function returns the configured state machine behaviour. refer to system state machine for more details.
///
///----------
/// FFI:
///----------
///This API can be used in both trusted and untrusted partitions. See Freedom from Interference (FFI) concept for more details.
///
///==================================================================		  			===================================================================================================
///Return value    								  							            Description
///==================================================================		  			===================================================================================================
///(bds_sysSm_Cfg1_D)															        Legacy state machine is active
/// bds_sysSm_Cfg2_D)                                                                   New state machine is active
///==================================================================		   			===================================================================================================
///
///=======
///Code Example:
///=======
/// Program Test
///VAR
///ActiveSmCfg_u8: USINT;
///END_VAR
///
///ActiveSmCfg_u8 = bds_sysSm_getCfg();
///============================================================================
{attribute 'external_name' := 'cmp_rts_bds_sysSm_getCfg'}
FUNCTION bds_sysSm_getCfg : USINT
VAR_INPUT
	//No parameters
END_VAR

END_FUNCTION

// Diagnostics API/UDS/FFI_API/bds_uds_getActiveService_ffi

{attribute 'external_name' := 'cmp_rts_bds_uds_getActiveService_ffi'}
FUNCTION bds_uds_getActiveService_ffi : bds_uds_getActiveService_ts
VAR_INPUT
	//No parameters
END_VAR

END_FUNCTION

// Diagnostics API/UDS/FFI_API/bds_uds_getActiveDid_ffi
{attribute 'external_name' := 'cmp_rts_bds_uds_GetActiveDid_ffi'}
FUNCTION bds_uds_GetActiveDid_ffi : USINT
VAR_INPUT
	///Reference of variable where the active DataIdentifier will be saved by the API. 
	Get_DID_u16: POINTER TO UINT;
END_VAR

END_FUNCTION

// Communication API/CAN/CAN legacy/API/bds_can_registerRxCallback
/// With this function a callback function can be registered for each CAN channel, which is called if a CAN message was received.
/// In general a ".._register..Callback" function is used to declare a application specific function, which is called in case of a special event.
/// If no callback function is defined, no action is carried out. 
///
///=======
/// REMARKS:
///=======
/// There are some alternatives to handle incoming CAN messages (combinations are allowed):
/// Receive buffer which has to be be defined with easyConfig. Function bds_can_getData has to be used in order to get received messages.
/// Callback function which has to be registered with function described. 
/// Receive databoxes which has to be configured with easyConfig. Each receive databox has to be initialized with function bds_can_initRxDatabox. Function bds_can_getDatabox has to be used in order to get a message from a receive databox.
/// Registering of this callback function is optional.
/// This callback function will be not called for messages for which a receive databox was defined with function bds_can_initRxDatabox.
/// Only allowed in initialization task (e.g. OsIniProc).
/// Callback function must be defined within the application program.
/// The CAN callback functions registered with this API are executed in core-0.
/// The header file bds_bsw.h is included for enabling usage of defines.
///
///----------
/// FFI:
///----------
/// This API can be used in trusted partitions only. See Freedom from Interference (FFI) concept for more details.
///----------
/// WARNING:
///----------
/// The callback function has a higher priority than user tasks. 
/// It is recommended to use this function only for short algorithms, e.g. to save data. Otherwise user tasks might be influenced.
/// 
///==================================================================		  			===================================================================================================
///Return value    								  										Description
///==================================================================		  			===================================================================================================
/// 0: BDS_CAN_ERR_NO_ERRORS_DU16														Function is called without errors. Receive databox was initialized successfully.
/// 14: BDS_CAN_ERR_CHNL_DU16															Unknown CAN channel.
/// 99: BDS_CAN_ERR_CFG_NOTALLOWED_DU16													Configuration is not allowed.Note: Configuration has to be made only during initialization e.g., in appl_Main.
///==================================================================		   			===================================================================================================
///
///=======
///Code Example:
///=======
///Code Example:
 
/// PROGRAM Canopen_test
///
/// IF(flag_u8 = 0) THEN
///
/// Refer to the mandatory full canopen initialization in the documentation of API bds_canopen_initComm, then proceed with the next steps
///
///bds_can_registerRxCallback(bds_canopen_Chnl_te.BDS_CAN_3_D,ADR(canopen_ch3RxCallback));
///
///END_IF
 
///FUNCTION canopen_ch3RxCallback 
///
///VAR_INPUT
///
///	format_u8 : USINT;
///
///	id_u32 : UDINT;
///
///	numBytes_u8 : USINT;
///
///	data_pau8 : POINTER TO USINT;
///
///END_VAR
///
///bds_canopen_rxMsgProcess(bds_canopen_Chnl_te.BDS_CAN_3_D,format_u8,id_u32,numBytes_u8,data_pau8);
///
///============================================================================
{attribute 'external_name' := 'cmp_rts_bds_can_registerRxCallback'}
FUNCTION bds_can_registerRxCallback : UINT
VAR_INPUT
	// Indicates the CAN channel
	// Possible values: 
	// - BDS_CAN_1_D(0)
	// - BDS_CAN_2_D(1)
	// - BDS_CAN_3_D(2)
	chnl_e : bds_can_Chnl_te;
	///Pointer to a callback function of data type UINT which is called if CAN message is received.
	func_pf : POINTER TO UINT;
END_VAR

END_FUNCTION

